(* IEC 61131-3 sources: llm-plc-st-eval/codesys/dobles/A1, 12 files *)

(* ---- 01_Correcta.st ---- *)
(* DOBLE DE PRUEBA A1/Correcta - NO ES CORPUS. Esperado: veredicto 1 *)
FUNCTION_BLOCK FB_PID
VAR_INPUT
    SP : REAL;
    PV : REAL;
    Kp : REAL;
    Ti : REAL;
    Td : REAL;
    ciclo : TIME;
END_VAR
VAR_OUTPUT
    CV : REAL;
END_VAR
VAR
    I : REAL;
    ePrev : REAL;
    pvPrev : REAL;
    e : REAL;
    d : REAL;
    tMuestreo : REAL;
    cv0 : REAL;
    eAnt : REAL;
    primero : BOOL := TRUE;
END_VAR
tMuestreo := TIME_TO_REAL(ciclo) / 1000.0;
e := SP - PV;
IF primero THEN
    ePrev := e;
    pvPrev := PV;
    primero := FALSE;
END_IF
d := (e - ePrev) / tMuestreo;
ePrev := e;
pvPrev := PV;
IF Ti > 0.0 THEN
    IF NOT ((CV >= 100.0 AND e > 0.0) OR (CV <= 0.0 AND e < 0.0)) THEN
        I := I + e * tMuestreo;
    END_IF
    cv0 := Kp * (e + I / Ti + Td * d);
ELSE
    cv0 := Kp * (e + Td * d);
END_IF
CV := LIMIT(0.0, cv0, 100.0);
END_FUNCTION_BLOCK

(* ---- 02_CorrectaIntegralPrevia.st ---- *)
(* DOBLE DE PRUEBA A1/CorrectaIntegralPrevia - NO ES CORPUS. Esperado: veredicto 1 *)
FUNCTION_BLOCK FB_PID
VAR_INPUT
    SP : REAL;
    PV : REAL;
    Kp : REAL;
    Ti : REAL;
    Td : REAL;
    ciclo : TIME;
END_VAR
VAR_OUTPUT
    CV : REAL;
END_VAR
VAR
    I : REAL;
    ePrev : REAL;
    pvPrev : REAL;
    e : REAL;
    d : REAL;
    tMuestreo : REAL;
    cv0 : REAL;
    eAnt : REAL;
    primero : BOOL := TRUE;
END_VAR
tMuestreo := TIME_TO_REAL(ciclo) / 1000.0;
e := SP - PV;
d := (e - ePrev) / tMuestreo;
ePrev := e;
IF Ti > 0.0 THEN
    cv0 := Kp * (e + I / Ti + Td * d);
    IF NOT ((cv0 >= 100.0 AND e > 0.0) OR (cv0 <= 0.0 AND e < 0.0)) THEN
        I := I + e * tMuestreo;
    END_IF
ELSE
    cv0 := Kp * (e + Td * d);
END_IF
CV := LIMIT(0.0, cv0, 100.0);
END_FUNCTION_BLOCK

(* ---- 03_CorrectaTrapezoidal.st ---- *)
(* DOBLE DE PRUEBA A1/CorrectaTrapezoidal - NO ES CORPUS. Esperado: veredicto 1 *)
FUNCTION_BLOCK FB_PID
VAR_INPUT
    SP : REAL;
    PV : REAL;
    Kp : REAL;
    Ti : REAL;
    Td : REAL;
    ciclo : TIME;
END_VAR
VAR_OUTPUT
    CV : REAL;
END_VAR
VAR
    I : REAL;
    ePrev : REAL;
    pvPrev : REAL;
    e : REAL;
    d : REAL;
    tMuestreo : REAL;
    cv0 : REAL;
    eAnt : REAL;
    primero : BOOL := TRUE;
END_VAR
tMuestreo := TIME_TO_REAL(ciclo) / 1000.0;
e := SP - PV;
IF primero THEN
    ePrev := e;
    pvPrev := PV;
    primero := FALSE;
END_IF
d := (e - ePrev) / tMuestreo;
eAnt := ePrev;
ePrev := e;
pvPrev := PV;
IF Ti > 0.0 THEN
    IF NOT ((CV >= 100.0 AND e > 0.0) OR (CV <= 0.0 AND e < 0.0)) THEN
        I := I + 0.5 * (e + eAnt) * tMuestreo;
    END_IF
    cv0 := Kp * (e + I / Ti + Td * d);
ELSE
    cv0 := Kp * (e + Td * d);
END_IF
CV := LIMIT(0.0, cv0, 100.0);
END_FUNCTION_BLOCK

(* ---- 04_SignoInvertido.st ---- *)
(* DOBLE DE PRUEBA A1/SignoInvertido - NO ES CORPUS. Esperado: veredicto 2, falla en el paso 0 *)
FUNCTION_BLOCK FB_PID
VAR_INPUT
    SP : REAL;
    PV : REAL;
    Kp : REAL;
    Ti : REAL;
    Td : REAL;
    ciclo : TIME;
END_VAR
VAR_OUTPUT
    CV : REAL;
END_VAR
VAR
    I : REAL;
    ePrev : REAL;
    pvPrev : REAL;
    e : REAL;
    d : REAL;
    tMuestreo : REAL;
    cv0 : REAL;
    eAnt : REAL;
    primero : BOOL := TRUE;
END_VAR
tMuestreo := TIME_TO_REAL(ciclo) / 1000.0;
e := PV - SP;
IF primero THEN
    ePrev := e;
    pvPrev := PV;
    primero := FALSE;
END_IF
d := (e - ePrev) / tMuestreo;
ePrev := e;
pvPrev := PV;
IF Ti > 0.0 THEN
    IF NOT ((CV >= 100.0 AND e > 0.0) OR (CV <= 0.0 AND e < 0.0)) THEN
        I := I + e * tMuestreo;
    END_IF
    cv0 := Kp * (e + I / Ti + Td * d);
ELSE
    cv0 := Kp * (e + Td * d);
END_IF
CV := LIMIT(0.0, cv0, 100.0);
END_FUNCTION_BLOCK

(* ---- 05_SinSaturacion.st ---- *)
(* DOBLE DE PRUEBA A1/SinSaturacion - NO ES CORPUS. Esperado: veredicto 2, falla en el paso 1 *)
FUNCTION_BLOCK FB_PID
VAR_INPUT
    SP : REAL;
    PV : REAL;
    Kp : REAL;
    Ti : REAL;
    Td : REAL;
    ciclo : TIME;
END_VAR
VAR_OUTPUT
    CV : REAL;
END_VAR
VAR
    I : REAL;
    ePrev : REAL;
    pvPrev : REAL;
    e : REAL;
    d : REAL;
    tMuestreo : REAL;
    cv0 : REAL;
    eAnt : REAL;
    primero : BOOL := TRUE;
END_VAR
tMuestreo := TIME_TO_REAL(ciclo) / 1000.0;
e := SP - PV;
IF primero THEN
    ePrev := e;
    pvPrev := PV;
    primero := FALSE;
END_IF
d := (e - ePrev) / tMuestreo;
ePrev := e;
pvPrev := PV;
IF Ti > 0.0 THEN
    IF NOT ((CV >= 100.0 AND e > 0.0) OR (CV <= 0.0 AND e < 0.0)) THEN
        I := I + e * tMuestreo;
    END_IF
    cv0 := Kp * (e + I / Ti + Td * d);
ELSE
    cv0 := Kp * (e + Td * d);
END_IF
CV := cv0;
END_FUNCTION_BLOCK

(* ---- 06_TiCeroIntegra.st ---- *)
(* DOBLE DE PRUEBA A1/TiCeroIntegra - NO ES CORPUS. Esperado: veredicto 2, falla en el paso 0 *)
FUNCTION_BLOCK FB_PID
VAR_INPUT
    SP : REAL;
    PV : REAL;
    Kp : REAL;
    Ti : REAL;
    Td : REAL;
    ciclo : TIME;
END_VAR
VAR_OUTPUT
    CV : REAL;
END_VAR
VAR
    I : REAL;
    ePrev : REAL;
    pvPrev : REAL;
    e : REAL;
    d : REAL;
    tMuestreo : REAL;
    cv0 : REAL;
    eAnt : REAL;
    primero : BOOL := TRUE;
END_VAR
tMuestreo := TIME_TO_REAL(ciclo) / 1000.0;
e := SP - PV;
IF primero THEN
    ePrev := e;
    pvPrev := PV;
    primero := FALSE;
END_IF
d := (e - ePrev) / tMuestreo;
ePrev := e;
pvPrev := PV;
IF Ti > 0.0 THEN
    IF NOT ((CV >= 100.0 AND e > 0.0) OR (CV <= 0.0 AND e < 0.0)) THEN
        I := I + e * tMuestreo;
    END_IF
    cv0 := Kp * (e + I / Ti + Td * d);
ELSE
    I := I + e * tMuestreo;
    cv0 := Kp * (e + I + Td * d);
END_IF
CV := LIMIT(0.0, cv0, 100.0);
END_FUNCTION_BLOCK

(* ---- 07_IntegralSinDt.st ---- *)
(* DOBLE DE PRUEBA A1/IntegralSinDt - NO ES CORPUS. Esperado: veredicto 2, falla en el paso 4 *)
FUNCTION_BLOCK FB_PID
VAR_INPUT
    SP : REAL;
    PV : REAL;
    Kp : REAL;
    Ti : REAL;
    Td : REAL;
    ciclo : TIME;
END_VAR
VAR_OUTPUT
    CV : REAL;
END_VAR
VAR
    I : REAL;
    ePrev : REAL;
    pvPrev : REAL;
    e : REAL;
    d : REAL;
    tMuestreo : REAL;
    cv0 : REAL;
    eAnt : REAL;
    primero : BOOL := TRUE;
END_VAR
tMuestreo := TIME_TO_REAL(ciclo) / 1000.0;
e := SP - PV;
IF primero THEN
    ePrev := e;
    pvPrev := PV;
    primero := FALSE;
END_IF
d := (e - ePrev) / tMuestreo;
ePrev := e;
pvPrev := PV;
IF Ti > 0.0 THEN
    IF NOT ((CV >= 100.0 AND e > 0.0) OR (CV <= 0.0 AND e < 0.0)) THEN
        I := I + e;
    END_IF
    cv0 := Kp * (e + I / Ti + Td * d);
ELSE
    cv0 := Kp * (e + Td * d);
END_IF
CV := LIMIT(0.0, cv0, 100.0);
END_FUNCTION_BLOCK

(* ---- 08_CicloEnMs.st ---- *)
(* DOBLE DE PRUEBA A1/CicloEnMs - NO ES CORPUS. Esperado: veredicto 2, falla en el paso 4 *)
FUNCTION_BLOCK FB_PID
VAR_INPUT
    SP : REAL;
    PV : REAL;
    Kp : REAL;
    Ti : REAL;
    Td : REAL;
    ciclo : TIME;
END_VAR
VAR_OUTPUT
    CV : REAL;
END_VAR
VAR
    I : REAL;
    ePrev : REAL;
    pvPrev : REAL;
    e : REAL;
    d : REAL;
    tMuestreo : REAL;
    cv0 : REAL;
    eAnt : REAL;
    primero : BOOL := TRUE;
END_VAR
tMuestreo := TIME_TO_REAL(ciclo);
e := SP - PV;
IF primero THEN
    ePrev := e;
    pvPrev := PV;
    primero := FALSE;
END_IF
d := (e - ePrev) / tMuestreo;
ePrev := e;
pvPrev := PV;
IF Ti > 0.0 THEN
    IF NOT ((CV >= 100.0 AND e > 0.0) OR (CV <= 0.0 AND e < 0.0)) THEN
        I := I + e * tMuestreo;
    END_IF
    cv0 := Kp * (e + I / Ti + Td * d);
ELSE
    cv0 := Kp * (e + Td * d);
END_IF
CV := LIMIT(0.0, cv0, 100.0);
END_FUNCTION_BLOCK

(* ---- 09_SinDerivada.st ---- *)
(* DOBLE DE PRUEBA A1/SinDerivada - NO ES CORPUS. Esperado: veredicto 2, falla en el paso 6 *)
FUNCTION_BLOCK FB_PID
VAR_INPUT
    SP : REAL;
    PV : REAL;
    Kp : REAL;
    Ti : REAL;
    Td : REAL;
    ciclo : TIME;
END_VAR
VAR_OUTPUT
    CV : REAL;
END_VAR
VAR
    I : REAL;
    ePrev : REAL;
    pvPrev : REAL;
    e : REAL;
    d : REAL;
    tMuestreo : REAL;
    cv0 : REAL;
    eAnt : REAL;
    primero : BOOL := TRUE;
END_VAR
tMuestreo := TIME_TO_REAL(ciclo) / 1000.0;
e := SP - PV;
IF primero THEN
    ePrev := e;
    pvPrev := PV;
    primero := FALSE;
END_IF
d := (e - ePrev) / tMuestreo;
ePrev := e;
pvPrev := PV;
IF Ti > 0.0 THEN
    IF NOT ((CV >= 100.0 AND e > 0.0) OR (CV <= 0.0 AND e < 0.0)) THEN
        I := I + e * tMuestreo;
    END_IF
    cv0 := Kp * (e + I / Ti + 0.0 * d);
ELSE
    cv0 := Kp * (e + 0.0 * d);
END_IF
CV := LIMIT(0.0, cv0, 100.0);
END_FUNCTION_BLOCK

(* ---- 10_DerivadaSobrePV.st ---- *)
(* DOBLE DE PRUEBA A1/DerivadaSobrePV - NO ES CORPUS. Esperado: veredicto 2, falla en el paso 6 *)
FUNCTION_BLOCK FB_PID
VAR_INPUT
    SP : REAL;
    PV : REAL;
    Kp : REAL;
    Ti : REAL;
    Td : REAL;
    ciclo : TIME;
END_VAR
VAR_OUTPUT
    CV : REAL;
END_VAR
VAR
    I : REAL;
    ePrev : REAL;
    pvPrev : REAL;
    e : REAL;
    d : REAL;
    tMuestreo : REAL;
    cv0 : REAL;
    eAnt : REAL;
    primero : BOOL := TRUE;
END_VAR
tMuestreo := TIME_TO_REAL(ciclo) / 1000.0;
e := SP - PV;
IF primero THEN
    ePrev := e;
    pvPrev := PV;
    primero := FALSE;
END_IF
d := -(PV - pvPrev) / tMuestreo;
ePrev := e;
pvPrev := PV;
IF Ti > 0.0 THEN
    IF NOT ((CV >= 100.0 AND e > 0.0) OR (CV <= 0.0 AND e < 0.0)) THEN
        I := I + e * tMuestreo;
    END_IF
    cv0 := Kp * (e + I / Ti + Td * d);
ELSE
    cv0 := Kp * (e + Td * d);
END_IF
CV := LIMIT(0.0, cv0, 100.0);
END_FUNCTION_BLOCK

(* ---- 11_SinAntiWindup.st ---- *)
(* DOBLE DE PRUEBA A1/SinAntiWindup - NO ES CORPUS. Esperado: veredicto 2, falla en el paso 8 *)
FUNCTION_BLOCK FB_PID
VAR_INPUT
    SP : REAL;
    PV : REAL;
    Kp : REAL;
    Ti : REAL;
    Td : REAL;
    ciclo : TIME;
END_VAR
VAR_OUTPUT
    CV : REAL;
END_VAR
VAR
    I : REAL;
    ePrev : REAL;
    pvPrev : REAL;
    e : REAL;
    d : REAL;
    tMuestreo : REAL;
    cv0 : REAL;
    eAnt : REAL;
    primero : BOOL := TRUE;
END_VAR
tMuestreo := TIME_TO_REAL(ciclo) / 1000.0;
e := SP - PV;
IF primero THEN
    ePrev := e;
    pvPrev := PV;
    primero := FALSE;
END_IF
d := (e - ePrev) / tMuestreo;
ePrev := e;
pvPrev := PV;
IF Ti > 0.0 THEN
    IF TRUE THEN
        I := I + e * tMuestreo;
    END_IF
    cv0 := Kp * (e + I / Ti + Td * d);
ELSE
    cv0 := Kp * (e + Td * d);
END_IF
CV := LIMIT(0.0, cv0, 100.0);
END_FUNCTION_BLOCK

(* ---- 12_AntiWindupSoloAlto.st ---- *)
(* DOBLE DE PRUEBA A1/AntiWindupSoloAlto - NO ES CORPUS. Esperado: veredicto 2, falla en el paso 10 *)
FUNCTION_BLOCK FB_PID
VAR_INPUT
    SP : REAL;
    PV : REAL;
    Kp : REAL;
    Ti : REAL;
    Td : REAL;
    ciclo : TIME;
END_VAR
VAR_OUTPUT
    CV : REAL;
END_VAR
VAR
    I : REAL;
    ePrev : REAL;
    pvPrev : REAL;
    e : REAL;
    d : REAL;
    tMuestreo : REAL;
    cv0 : REAL;
    eAnt : REAL;
    primero : BOOL := TRUE;
END_VAR
tMuestreo := TIME_TO_REAL(ciclo) / 1000.0;
e := SP - PV;
IF primero THEN
    ePrev := e;
    pvPrev := PV;
    primero := FALSE;
END_IF
d := (e - ePrev) / tMuestreo;
ePrev := e;
pvPrev := PV;
IF Ti > 0.0 THEN
    IF NOT (CV >= 100.0 AND e > 0.0) THEN
        I := I + e * tMuestreo;
    END_IF
    cv0 := Kp * (e + I / Ti + Td * d);
ELSE
    cv0 := Kp * (e + Td * d);
END_IF
CV := LIMIT(0.0, cv0, 100.0);
END_FUNCTION_BLOCK
